SUBAPPLICATION TimedFunc (* Subapplication Type *)
  (* Standard: 61499-2 *)
  (* Version 1.0, 2023-01-29, Franz *)
  IMPORT isobus::UT::io::Softkey::SoftKeyActivationCode::SK_RELEASED;
  IMPORT isobus::UT::io::Auxiliary::IN::AuxiliaryState::AuxDisabled;
  IMPORT logiBUS::io::DQ::logiBUS_DO::Invalid;
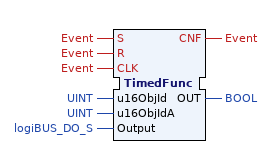
  EVENT_INPUT
    S; (* Set output Q *)
    R; (* Reset output Q *)
    CLK; (* Clock for triggering a output toggle *)
  END_EVENT
  EVENT_OUTPUT
    CNF;
  END_EVENT
  VAR_INPUT
    u16ObjId : UINT;
    u16ObjIdA : UINT;
    Output : logiBUS::io::DQ::logiBUS_DO_S := Invalid;
  END_VAR
  VAR_OUTPUT
    OUT : BOOL;
  END_VAR
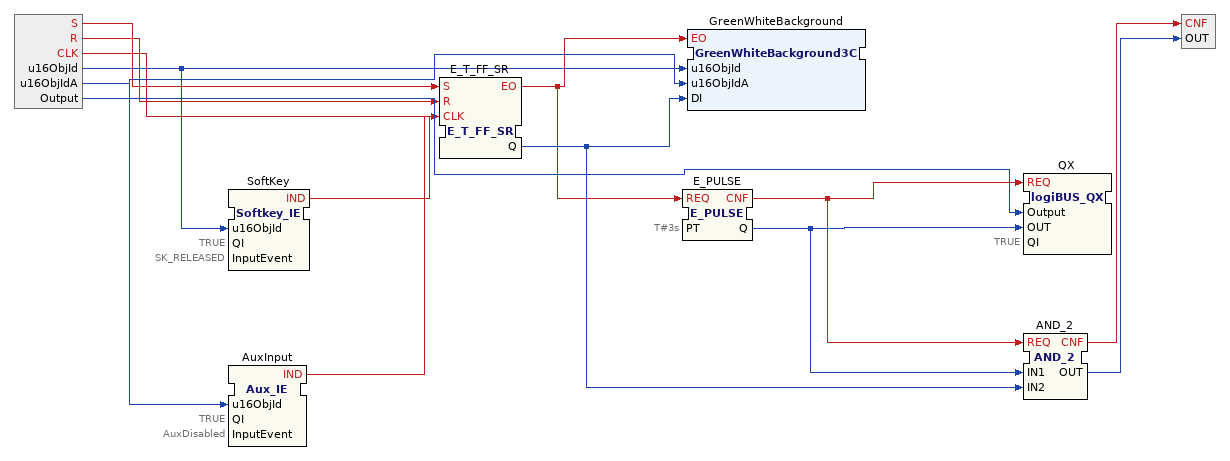
  FBS
    AND_2 : iec61131::bitwiseOperators::AND_2;
    QX : logiBUS::io::DQ::logiBUS_QX(QI := TRUE);
    E_PULSE : iec61499::events::timers::E_PULSE(PT := T#3s);
    E_T_FF_SR : iec61499::events::E_T_FF_SR;
    SoftKey : isobus::UT::io::Softkey::Softkey_IE(QI := TRUE, InputEvent := SK_RELEASED);
    AuxInput : isobus::UT::io::Auxiliary::IN::Aux_IE(QI := TRUE, InputEvent := AuxDisabled);
  END_FBS
  SUBAPPS
    GreenWhiteBackground : MyLib::sys::GreenWhiteBackground3C;
  END_SUBAPPS
  EVENT_CONNECTIONS
    E_PULSE.CNF TO AND_2.REQ;
    E_PULSE.CNF TO QX.REQ;
    AND_2.CNF TO CNF;
    E_T_FF_SR.EO TO E_PULSE.REQ;
    E_T_FF_SR.EO TO GreenWhiteBackground.EO;
    S TO E_T_FF_SR.S;
    R TO E_T_FF_SR.R;
    CLK TO E_T_FF_SR.CLK;
    SoftKey.IND TO E_T_FF_SR.CLK;
    AuxInput.IND TO E_T_FF_SR.CLK;
  END_CONNECTIONS
  DATA_CONNECTIONS
    Output TO QX.Output;
    u16ObjIdA TO AuxInput.u16ObjId;
    u16ObjId TO SoftKey.u16ObjId;
    AND_2.OUT TO OUT;
    u16ObjId TO GreenWhiteBackground.u16ObjId;
    u16ObjIdA TO GreenWhiteBackground.u16ObjIdA;
    E_PULSE.Q TO QX.OUT;
    E_PULSE.Q TO AND_2.IN1;
    E_T_FF_SR.Q TO AND_2.IN2;
    E_T_FF_SR.Q TO GreenWhiteBackground.DI;
  END_CONNECTIONS
END_SUBAPPLICATION
